Fanuc KAREL source: KA00103.KL

PROGRAM KA00103
%NOLOCKGROUP
VAR
  SRC: VECTOR
  DST: XYZWPREXT
BEGIN
  SRC.X = 1.0
  DST = SRC
END KA00103
